# EPICS substitutions: db/Beckhoff_7XXX/ecmcEP7211-0034_OPT_common.substitutions
# Actual torque is mapped in every OPT mode.
file "ecmc_analogInput-chX.template"
{
  pattern {CH_ID, sourceName, KEY, suffix, DESC, EGU, ESLO, PREC, LOPR, HOPR, LOLO, LOW, HIGH, HIHI, HYST, LLSV, LSV, HSV, HHSV}
          {01,    "torqueActual",   "Drv", "-TrqAct", "Actual Trq", "%",     0.1,       1,    -200, 200,  0,    -80, 80,   0,    0,    "NO_ALARM", "NO_ALARM", "MINOR",    "NO_ALARM"}
}
